(* CODESYS project GVL_Alarm.gvl.xml

Project tree, tasks and I/O mapping:
  global variables GVL_Alarm
*)

// GVL_Alarm
{attribute 'qualified_only'}
VAR_GLOBAL
	AlarmConstant : DINT := 3;
END_VAR
